(*
SPDX-FileCopyrightText: © 2026 Oleksandr Tiutyk <trofimich@gmail.com>
SPDX-License-Identifier: MIT
License: https://opensource.org/license/mit
*)

(*!
<summary>Resolves externally managed dependencies by a stable key.</summary>
<description>
Resolution borrows an existing shared instance without transferring ownership.
Return zero for an unknown key.
</description>
*)
INTERFACE IWorkflowDependencyResolver

(*!
<summary>Returns an existing borrowed dependency for the supplied stable key.</summary>
<description>Return zero for an unknown key.</description>
<param name="key">Dependency lookup key.</param>
*)
METHOD ResolveExternal : TOF_Core.IObject
VAR_INPUT
	key : STRING;
END_VAR
END_METHOD

END_INTERFACE

(* stored: Version 1.1.0.1
   Itf IWorkflowDependencyResolver: Id {b7b88fc9-3040-442b-8f55-f4771df1f971}
   Method ResolveExternal: Id {89234413-f41f-4f3e-9eae-ab747312db5a} *)
